Fanuc KAREL source: KT00515.KL

PROGRAM KT00515
%NOLOCKGROUP
VAR
  P1: XYZWPREXT
  P2: POSITION
  OUT: XYZWPR
BEGIN
  P1.X = 1.0
  OUT = P1 : P2
END KT00515
